(*
SPDX-FileCopyrightText: © 2026 Oleksandr Tiutyk <trofimich@gmail.com>
SPDX-License-Identifier: MIT
License: https://opensource.org/license/mit
*)

(*!
<summary>Names the operations and successful completion of DirectoryTest scenarios.</summary>
<description>
Each scenario follows its explicit subset of steps. Advancing requires the expected stop reason and any
existence checks for that step. COMPLETED ends scenario work. Cleanup advances on later test cycles.
The enum is internal to the tests.
</description>
*)
{attribute 'qualified_only'}
{attribute 'strict'}
{attribute 'to_string'}
TYPE DIRECTORY_TEST_STEP :
(
	//! <summary>Create the test directory; success establishes ownership, an existing path causes failure.</summary>
	CREATE_DIRECTORY := 0,
	//! <summary>Verify the newly created test directory exists.</summary>
	CHECK_DIRECTORY_PRESENT,
	//! <summary>Create a child directory inside the owned test directory.</summary>
	CREATE_CHILD_DIRECTORY,
	//! <summary>Verify the first conditional creation produced a child directory.</summary>
	CHECK_CHILD_DIRECTORY_PRESENT,
	//! <summary>Repeat conditional creation while the child directory exists.</summary>
	CREATE_CHILD_DIRECTORY_AGAIN,
	//! <summary>Verify the child directory still exists after repeated creation.</summary>
	CHECK_CHILD_DIRECTORY_PRESENT_AGAIN,
	//! <summary>Require native removal of the nonempty parent directory to fail.</summary>
	REJECT_NONEMPTY_DIRECTORY_REMOVAL,
	//! <summary>Confirm the child still exists after the failed parent removal.</summary>
	CHECK_CHILD_DIRECTORY_RETAINED,
	//! <summary>Remove the owned child directory using conditional removal.</summary>
	REMOVE_CHILD_DIRECTORY,
	//! <summary>Verify that the child directory is absent.</summary>
	CHECK_CHILD_DIRECTORY_ABSENT,
	//! <summary>Repeat conditional removal while the child directory is absent.</summary>
	REMOVE_CHILD_DIRECTORY_AGAIN,
	//! <summary>Verify the child directory is still absent after repeated removal.</summary>
	CHECK_CHILD_DIRECTORY_ABSENT_AGAIN,
	//! <summary>Remove the empty test directory created by this scenario.</summary>
	REMOVE_DIRECTORY,
	//! <summary>Verify the test directory is absent after removal.</summary>
	CHECK_DIRECTORY_ABSENT,
	//! <summary>All scenario operations and postconditions completed successfully.</summary>
	COMPLETED
);
END_TYPE

(* stored: Version 1.1.0.1
   DUT DIRECTORY_TEST_STEP: Id {bf4fd83d-636c-4583-83cd-68d10caca698} *)
